(* IEC 61131-3 sources: kns-pump-station/tests/POUs/Station/FB_StationAlarms_Test, 14 files *)

(* ---- AckAllViaInterface.method.decl.st ---- *)
// PL.I_AlarmSource.AckAll (сводка, общий сброс): квитирует все тревоги станции ближайшим вызовом
METHOD PRIVATE AckAllViaInterface
VAR
    fbDut  : FB_StationAlarms;          // ФБ под тестом
    fbTime : PL.FB_FakeTime;            // подменное время, старт 1 ч
    stCfg  : ST_StationCfg;             // тревоги по умолчанию (05_alarm_list.csv)
    itfSrc : PL.I_AlarmSource;        // источник через интерфейс
END_VAR

(* ---- AckMaskAcksSlot.method.decl.st ---- *)
// 04 §19.2: маска wAckReq, бит slot - 1, квитирует свою тревогу, остальные — нет
METHOD PRIVATE AckMaskAcksSlot
VAR
    fbDut  : FB_StationAlarms;          // ФБ под тестом
    fbTime : PL.FB_FakeTime;            // подменное время, старт 1 ч
    stCfg  : ST_StationCfg;             // тревоги по умолчанию (05_alarm_list.csv)
    itfAlm : PL.I_Alarm;              // тревога через интерфейс
END_VAR

(* ---- GetAlarmIndexOutOfRangeReturnsZero.method.decl.st ---- *)
// PL.I_AlarmSource.GetAlarm вне 0…AlarmCount - 1 — 0
METHOD PRIVATE GetAlarmIndexOutOfRangeReturnsZero
VAR
    fbDut  : FB_StationAlarms;          // ФБ под тестом
    fbTime : PL.FB_FakeTime;            // подменное время, старт 1 ч
    stCfg  : ST_StationCfg;             // тревоги по умолчанию (05_alarm_list.csv)
    itfAlm : PL.I_Alarm;              // тревога через интерфейс
END_VAR

(* ---- IdsAreBasePlusSlot.method.decl.st ---- *)
// 04 §15, API 20.5: номер тревоги = 100000 + slot; индекс источника 0 — slot 1; AlarmCount = 13
METHOD PRIVATE IdsAreBasePlusSlot
VAR
    fbDut  : FB_StationAlarms;          // ФБ под тестом
    fbTime : PL.FB_FakeTime;            // подменное время, старт 1 ч
    stCfg  : ST_StationCfg;             // тревоги по умолчанию (05_alarm_list.csv)
    itfAlm : PL.I_Alarm;              // тревога через интерфейс
    uiIdx  : UINT;                    // индекс источника
    xIdsOk : BOOL := TRUE;            // все номера верны
END_VAR

(* ---- IdsAreBasePlusSlot.method.impl.st ---- *)
coUnit.TEST('StationAlarms_IdsAreBasePlusSlot_A15');

fbDut(itfTime := fbTime, stCfg := stCfg);
AssertEquals_UINT(Expected := 13, Actual := fbDut.AlarmCount, Message := '13 station alarms');
FOR uiIdx := 0 TO 12 DO
    itfAlm := fbDut.GetAlarm(uiIndex := uiIdx);
    IF itfAlm = 0 THEN
        xIdsOk := FALSE;
    ELSIF itfAlm.Id <> 100001 + UINT_TO_UDINT(uiIdx) THEN
        xIdsOk := FALSE;
    END_IF
END_FOR
AssertTrue(Condition := xIdsOk, Message := 'ids 100001...100013');
itfAlm := fbDut.GetAlarm(uiIndex := E_StationAlarm.ATS - 1);
AssertEquals_UDINT(Expected := 100005, Actual := itfAlm.Id, Message := 'KNS1.ATS = 100005');

coUnit.TEST_FINISHED();

(* ---- OnDelayFromCfg.method.decl.st ---- *)
// 05_alarm_list.csv: задержка появления KNS1.LACK 10 с — из Cfg тревоги (не раньше)
METHOD PRIVATE OnDelayFromCfg
VAR
    fbDut  : FB_StationAlarms;          // ФБ под тестом
    fbTime : PL.FB_FakeTime;            // подменное время, старт 1 ч
    stCfg  : ST_StationCfg;             // тревоги по умолчанию (05_alarm_list.csv)
    uiStep : UINT;                    // шаг 100 мс
END_VAR

(* ---- OnDelayFromCfg.method.impl.st ---- *)
coUnit.TEST('StationAlarms_OnDelayFromCfg_A15_PMI17');

fbDut.axCond[E_StationAlarm.LACK] := TRUE;
fbDut(itfTime := fbTime, stCfg := stCfg);
FOR uiStep := 1 TO 99 DO
    fbTime.Advance(tStep := T#100MS);
    fbDut(itfTime := fbTime, stCfg := stCfg);
END_FOR
AssertEquals_WORD(Expected := 0, Actual := fbDut.wAlmActive, Message := 'LACK not active at 9.9 s');
fbTime.Advance(tStep := T#100MS);
fbDut(itfTime := fbTime, stCfg := stCfg);
AssertEquals_WORD(Expected := 16#0004, Actual := fbDut.wAlmActive, Message := 'LACK active at 10 s');

coUnit.TEST_FINISHED();

(* ---- ShelveRejectedForEhl.method.decl.st ---- *)
// 04 §15, PMI-36 шаг 6: KNS1.EHL отложить нельзя (tShelveMax = 0); DRY откладывается и возвращается масками
METHOD PRIVATE ShelveRejectedForEhl
VAR
    fbDut  : FB_StationAlarms;          // ФБ под тестом
    fbTime : PL.FB_FakeTime;            // подменное время, старт 1 ч
    stCfg  : ST_StationCfg;             // тревоги по умолчанию (05_alarm_list.csv)
    itfAlm : PL.I_Alarm;              // тревога через интерфейс
END_VAR

(* ---- SuppressionPutsSuppressedByDesign.method.decl.st ---- *)
// 04 §15, PMI-21: подавление по условию — SuppressedByDesign без неквитированности, бит в wAlmShelved
METHOD PRIVATE SuppressionPutsSuppressedByDesign
VAR
    fbDut  : FB_StationAlarms;          // ФБ под тестом
    fbTime : PL.FB_FakeTime;            // подменное время, старт 1 ч
    stCfg  : ST_StationCfg;             // тревоги по умолчанию (05_alarm_list.csv)
    itfAlm : PL.I_Alarm;              // тревога через интерфейс
END_VAR

(* ---- SuppressionReleaseRestartsOnDelay.method.decl.st ---- *)
// 04 §15, PMI-22, PMI-34: подавление по условию снято, а условие держится ещё цикл (станция видит выходы устройств
// циклом позже: после снятия «сухого хода» или восстановления питания насосы ещё «недоступны») — тревога не
// появляется: выдержка появления отсчитывается заново после снятия подавления (без мелькания High с сиреной)
METHOD PRIVATE SuppressionReleaseRestartsOnDelay
VAR
    fbDut  : FB_StationAlarms;          // ФБ под тестом
    fbTime : PL.FB_FakeTime;            // подменное время, старт 1 ч
    stCfg  : ST_StationCfg;             // тревоги по умолчанию (05_alarm_list.csv): NORES — 10 с
    itfAlm : PL.I_Alarm;                // тревога через интерфейс
    uiStep : UINT;                      // шаг времени
END_VAR

(* ---- SuppressionReleaseRestartsOnDelay.method.impl.st ---- *)
coUnit.TEST('StationAlarms_SuppressionReleaseRestartsOnDelay_A15_PMI22_PMI34');

fbDut.axCond[E_StationAlarm.NORES] := TRUE;
fbDut.axSuppress[E_StationAlarm.NORES] := TRUE;
FOR uiStep := 1 TO 150 DO
    fbTime.Advance(tStep := T#100MS);
    fbDut(itfTime := fbTime, stCfg := stCfg);
END_FOR
itfAlm := fbDut.GetAlarm(uiIndex := E_StationAlarm.NORES - 1);
AssertTrue(Condition := itfAlm.State = PL.E_AlarmState.SuppressedByDesign, Message := 'NORES suppressed for 15 s');
fbDut.axSuppress[E_StationAlarm.NORES] := FALSE;
fbTime.Advance(tStep := T#100MS);
fbDut(itfTime := fbTime, stCfg := stCfg);
AssertEquals_WORD(Expected := 0, Actual := fbDut.wAlmUnack, Message := 'no unacked alarm on suppression release');
AssertTrue(Condition := itfAlm.State = PL.E_AlarmState.Normal, Message := 'NORES normal right after release');
fbDut.axCond[E_StationAlarm.NORES] := FALSE;
fbTime.Advance(tStep := T#100MS);
fbDut(itfTime := fbTime, stCfg := stCfg);
AssertEquals_WORD(Expected := 0, Actual := fbDut.wAlmUnack, Message := 'nothing to acknowledge');
AssertTrue(Condition := fbDut.ePrioUnack = PL.E_AlarmPriority.None, Message := 'no unacked priority (no siren)');
// условие держится после снятия подавления — тревога через свою выдержку 10 с
fbDut.axCond[E_StationAlarm.NORES] := TRUE;
fbDut(itfTime := fbTime, stCfg := stCfg);
FOR uiStep := 1 TO 99 DO
    fbTime.Advance(tStep := T#100MS);
    fbDut(itfTime := fbTime, stCfg := stCfg);
END_FOR
AssertTrue(Condition := itfAlm.State = PL.E_AlarmState.Normal, Message := 'still normal at 9.9 s');
fbTime.Advance(tStep := T#100MS);
fbDut(itfTime := fbTime, stCfg := stCfg);
AssertTrue(Condition := itfAlm.State = PL.E_AlarmState.ActiveUnack, Message := 'NORES after its 10 s delay');

coUnit.TEST_FINISHED();

(* ---- TimeBackwardsOnDelayRestarts.method.decl.st ---- *)
// Время назад — задержка появления тревоги из Cfg отсчитывается заново
METHOD PRIVATE TimeBackwardsOnDelayRestarts
VAR
    fbDut  : FB_StationAlarms;          // ФБ под тестом
    fbTime : PL.FB_FakeTime;            // подменное время, старт 1 ч
    stCfg  : ST_StationCfg;             // тревоги по умолчанию (05_alarm_list.csv)
    uiStep : UINT;                    // шаг 100 мс
END_VAR

(* ---- TimeBackwardsOnDelayRestarts.method.impl.st ---- *)
coUnit.TEST('StationAlarms_TimeBackwardsOnDelayRestarts_A15');

fbDut.axCond[E_StationAlarm.LACK] := TRUE;
fbDut(itfTime := fbTime, stCfg := stCfg);
fbTime.Advance(tStep := T#5S);
fbDut(itfTime := fbTime, stCfg := stCfg);
fbTime.SetNow(ltValue := LTIME#59M);
FOR uiStep := 1 TO 100 DO
    fbTime.Advance(tStep := T#100MS);
    fbDut(itfTime := fbTime, stCfg := stCfg);
END_FOR
AssertEquals_WORD(Expected := 0, Actual := fbDut.wAlmActive, Message := 'on-delay restarted after time jump');
fbTime.Advance(tStep := T#100MS);
fbDut(itfTime := fbTime, stCfg := stCfg);
AssertEquals_WORD(Expected := 16#0004, Actual := fbDut.wAlmActive, Message := 'active after full on-delay');

coUnit.TEST_FINISHED();

(* ---- WordsAndPrioUnack.method.decl.st ---- *)
// 04 §19.3: слова wAlmActive, wAlmUnack и высший приоритет неквитированных (Critical EHL выше Low SIM)
METHOD PRIVATE WordsAndPrioUnack
VAR
    fbDut  : FB_StationAlarms;          // ФБ под тестом
    fbTime : PL.FB_FakeTime;            // подменное время, старт 1 ч
    stCfg  : ST_StationCfg;             // тревоги по умолчанию (05_alarm_list.csv)
END_VAR
